Fanuc KAREL source: kb00188.KL

-- PROVISIONAL review KL for V770-1; original PC SHA256 99db196e0dbe6b32a8723578ab9c84d11e255b56594e203c6f8cfb1a3258d489
-- Incomplete behavior may be omitted. Consult companion uncertainty JSON. Do not deploy.
PROGRAM KB00188
%NOLOCKGROUP
VAR
  P1 : STRING[80]
  RESULT : INTEGER
BEGIN
  -- UNRESOLVED_PC offsets 5-14; opcodes 3F,75
  -- UNRESOLVED_PC offsets 19-36; opcodes 27,22,2A,76,23
  -- UNRESOLVED_PC offsets 41-45; opcodes 7F
END KB00188
